TYPE ST_SwitchControlInput :
STRUCT
    nSwitchId      : UINT;
    stControlData  : ST_SwitchControlData;
END_STRUCT
END_TYPE

(* stored: Version 1.1.0.1, ProductVersion 3.1.4026.20
   DUT ST_SwitchControlInput: Id {D1A10004-0A11-4A11-8A11-000000000004} *)
